// TIA Portal V20 export
// export: Created 2026-10-20T12:52:53.0506322Z, ExportSetting WithDefaults, DisplayName Totally Integrated Automation Portal, DisplayVersion V20 Update 6, DisplayName TIA Portal Openness, DisplayVersion V20 Update 6, DisplayName TIA Portal Version Control Interface, DisplayVersion V20 Update 6, DisplayName SINAMICS Startdrive Advanced, DisplayVersion V20 SP1, DisplayName SINAMICS Startdrive G130, G150, S120, S150, SINAMICS MV, G220, S200, S210, DisplayVersion V20 SP1, DisplayName SINAMICS Startdrive G110M, G120, G120C, G120D, G120P, G115D, DisplayVersion V20 SP1, DisplayName STEP 7 Professional, DisplayVersion V20 Update 6, DisplayName STEP 7 Safety, DisplayVersion V20 Update 2, DisplayName WinCC Basic/Comfort/Advanced, DisplayVersion V20 Update 6, DisplayName WinCC Unified, DisplayVersion V20 Update 6
FUNCTION "Handshake_Infeed_FC" : Void   // FC47, SCL
{ S7_Optimized_Access := 'TRUE' }
VERSION : 0.1
// stored: AutoNumber true, IsIECCheckEnabled false, SetENOAutomatically false, UDAEnableTagReadback false
   VAR_INPUT
      Infeed_Stop_Sensor : Bool;
      Ready_To_Receive : Bool;
      Auto_Mode : Bool;
      Transfer_In_Progress : Bool;
      DB_LGX_To_SM_Infeed_Ready_To_Send : Bool;
      DB_LGX_To_SM_Infeed_Transfer_In_Progress : Bool;
   END_VAR
   VAR_OUTPUT
      Fault_Handshake : Bool;
      DB_SM_To_LGX_Infeed_Ready_To_Receive : Bool;
      DB_SM_To_LGX_Infeed_Pallet_Received : Bool;
      DB_SM_To_LGX_Infeed_Transfer_In_Progress : Bool;
   END_VAR
   VAR_TEMP
      tReady_To_Receive_Condition : Bool;
      tPallet_Received_Condition : Bool;
   END_VAR
BEGIN
   // ---------------------------------------------------------
   // STEP 1: Is SM ready to receive?
   // Condition: SM in Auto, infeed conveyor healthy,
   //            no transfer in progress, no alarm
   // ---------------------------------------------------------
   #tReady_To_Receive_Condition :=
   #Auto_Mode
   AND #Ready_To_Receive
   AND NOT #DB_SM_To_LGX_Infeed_Ready_To_Receive
   AND NOT #DB_SM_To_LGX_Infeed_Pallet_Received;

   IF #DB_LGX_To_SM_Infeed_Ready_To_Send
       AND #tReady_To_Receive_Condition THEN
       #DB_SM_To_LGX_Infeed_Ready_To_Receive := TRUE;
   END_IF;

   // ---------------------------------------------------------
   // STEP 2: Confirm pallet received
   // Condition: Photocell active while transfer is in progress
   // ---------------------------------------------------------
   // #tPallet_Received_Condition :=
   // #Infeed_Stop_Sensor
   // AND #DB_LGX_To_SM_Infeed_Transfer_In_Progress
   // AND #DB_SM_To_LGX_Infeed_Ready_To_Receive;
   // 
   #tPallet_Received_Condition :=
   #Infeed_Stop_Sensor;

   IF #tPallet_Received_Condition THEN
       #DB_SM_To_LGX_Infeed_Pallet_Received := TRUE;
       #DB_SM_To_LGX_Infeed_Ready_To_Receive := FALSE;
   ELSE
       #DB_SM_To_LGX_Infeed_Pallet_Received := FALSE;
   END_IF;

   // ---------------------------------------------------------
   // STEP 3: Reset after LGX confirms end of transfer
   // (LGX resets Transfer_In_Progress upon receiving Pallet_Received)
   // ---------------------------------------------------------
   // IF #DB_SM_To_LGX_Infeed_Pallet_Received
   //     AND NOT #DB_LGX_To_SM_Infeed_Transfer_In_Progress THEN
   //     #DB_SM_To_LGX_Infeed_Pallet_Received := FALSE;
   // END_IF;

   // ---------------------------------------------------------
   // STEP 4: Reset Ready_To_Receive if LGX withdraws Ready_To_Send
   // (e.g. LGX cancelled the operation before starting transfer)
   // ---------------------------------------------------------
   IF NOT #DB_LGX_To_SM_Infeed_Ready_To_Send
       AND NOT #DB_LGX_To_SM_Infeed_Transfer_In_Progress THEN
       #DB_SM_To_LGX_Infeed_Ready_To_Receive := FALSE;
   END_IF;

   // ---------------------------------------------------------
   // FAULT SUPERVISION
   // If Transfer_In_Progress remains active without pallet arriving:
   // use external timer / timeout bit (implement in OB1)
   // ---------------------------------------------------------
   #Fault_Handshake := FALSE; // Placeholder - implement watchdog

   #DB_SM_To_LGX_Infeed_Transfer_In_Progress := #Transfer_In_Progress;
END_FUNCTION
